// TIA Portal V21 export
// export: Created 2026-11-10T19:11:36.2534764Z, ExportSetting WithDefaults, DisplayName Totally Integrated Automation Portal, DisplayVersion V21 Update 3, DisplayName STEP 7 Professional, DisplayVersion V21 Update 3, DisplayName STEP 7 Safety, DisplayVersion V21, DisplayName Tech WebApplication, DisplayVersion V21, DisplayName WinCC Basic/Comfort/Advanced, DisplayVersion V21 Update 3, DisplayName WinCC Unified, DisplayVersion V21 Update 3
DATA_BLOCK "DB_SETIO_PART"   // DB20
// stored: AutoNumber true, DBAccessibleFromOPCUA true, DBAccessibleFromWebserver true, InstanceOfName SETIO_PART, OfSystemLibElement SETIO_PART, OfSystemLibVersion 1.2
"SETIO_PART"
   // VAR_INPUT
   //    ID : HW_SUBMODULE;
   //    OFFSET : Int;
   //    LEN : Int;
   // END_VAR
   // VAR_OUTPUT
   //    STATUS : DWord;
   //    ERROR : Bool;
   // END_VAR
   // VAR_IN_OUT
   //    OUTPUTS : Variant;
   // END_VAR
BEGIN
END_DATA_BLOCK
